Fanuc KAREL source: kb00018.compact.KL

PROGRAM KB00018
%STACKSIZE=65535
%PRIORITY=65535
%NOLOCKGROUP
VAR
P1 : XYZWPREXT
P2 : POSITION
P3 : POSITION
P4 : INTEGER
BEGIN
P4=1
CHECK_EPOS(P1,P2,P3,P4,1)
END KB00018
